Fanuc KAREL source: KX00029.KL

PROGRAM KX00029
%NOLOCKGROUP
%NOABORT = ERROR + COMMAND
VAR
  I: INTEGER
  J: INTEGER
  B: BOOLEAN
  F: FILE
  S: STRING[80]
  P: XYZWPR
BEGIN
  I = 1
END KX00029
